TYPE "ST_DeclarationUnitHal"
VERSION : 0.1
   STRUCT
      Cell { ExternalAccessible := 'False'; ExternalVisible := 'False'; ExternalWritable := 'False'} : "ST_DeclarationCellHal";
      Satellite { ExternalAccessible := 'False'; ExternalVisible := 'False'; ExternalWritable := 'False'} : "ST_SatelliteUnitHal";
   END_STRUCT;

END_TYPE

